RoboDK station: pick and place normal 2r.rdk

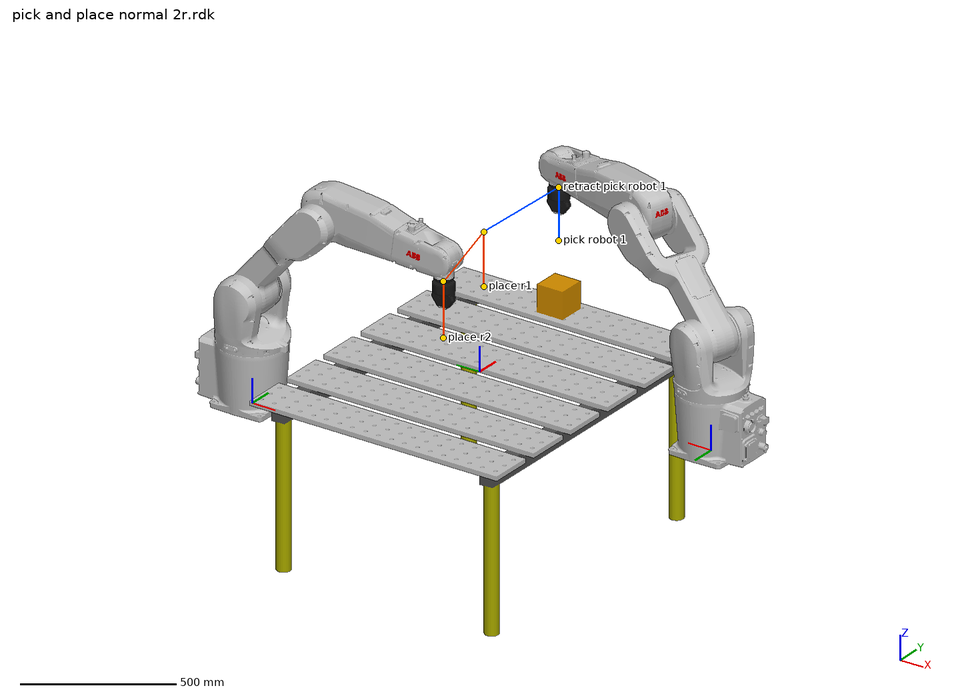
[picture v0: the station drawn from its stored meshes, robots at their saved joint values, targets as dots, program paths as lines]
Station pick and place normal 2r (saved by RoboDK 5.5.0). Poses are relative to the parent item; angles as X-Y-Z fixed-axis rotations.
  - frame Frame 2 at (700, 0, 200) mm, rotated rx 0 ry 0 rz 90 deg
    - object Table 1200x1000mm (Welding) at (0, 0, 0) mm, size 1193.8 x 965.2 x 609.6 mm, geometry from Table-1200x1000mm-Welding.sld
    - object Cube 100mm at (460, 0, 0) mm, size 100 x 100 x 100 mm, geometry from Cube-100mm.sld
  - frame ABB IRB 1200-5/0.9 (1) at (1400, 290, 0) mm, rotated rx 0 ry 0 rz 180 deg
    - robot ABB IRB 1200-5/0.9: 6 axes, payload 5 kg, reach 901 mm, repeatability 0.02 mm, weight 52 kg
        modified DH rows (alpha deg, a mm, theta deg, d mm): 0, 0, 0, 399; -90, 0, -90, 0; 0, 448, 0, 0; -90, 42, 0, 451; 90, 0, 0, 0; -90, 0, 180, 82
        joint limits [-170, -100, -200, -270, -130, -360] to [170, 130, 70, 270, 130, 360]; home [0, 0, 0, 0, 0, 0]; saved at [-16.36, 47.146, -44.021, 0, 86.875, -16.36]
      - robot RobotiQ 2F-140 Gripper (Mechanism) (model RobotiQ 2F140): 1 axes, payload 5 kg
          joint limits [0] to [140]; home [140]; saved at [140]
    - target pick robot 1 (Cartesian target) at (749.42, -220, 449.05) mm, rotated rx 180 ry 0 rz -180 deg; joints [-16.36, 51.781, -27.774, 0, 65.993, -16.36] of ABB IRB 1200-5/0.9
    - target retract pick robot 1 (Cartesian target) at (749.42, -220, 639.05) mm, rotated rx 180 ry 0 rz -180 deg; joints [-16.36, 47.146, -44.021, 0, 86.875, -16.36] of ABB IRB 1200-5/0.9
    - target retract place r1 (Cartesian target) at (759, 184.18, 639.12) mm, rotated rx 180 ry 0.01 rz -179.36 deg; joints [13.64, 47.14, -44.02, 0, 86.87, 13] of ABB IRB 1200-5/0.9
    - target place r1 (Cartesian target) at (759.03, 184.19, 444.12) mm, rotated rx 180 ry 0.01 rz -179.36 deg; joints [13.64, 52.024, -27.559, 0, 65.525, 13] of ABB IRB 1200-5/0.9
  - frame ABB IRB 1200-5/0.9 (2) at (0, -270, 0) mm
    - robot ABB IRB 1200-5/0.9: 6 axes, payload 5 kg, reach 901 mm, repeatability 0.02 mm, weight 52 kg
        modified DH rows (alpha deg, a mm, theta deg, d mm): 0, 0, 0, 399; -90, 0, -90, 0; 0, 448, 0, 0; -90, 42, 0, 451; 90, 0, 0, 0; -90, 0, 180, 82
        joint limits [-170, -100, -200, -270, -130, -360] to [170, 130, 70, 270, 130, 360]; home [0, 0, 0, 0, 0, 0]; saved at [0.38, 40.43, -32.71, 0, 82.29, -180.25]
      - robot RobotiQ 2F-140 Gripper (Mechanism) (model RobotiQ 2F140): 1 axes, payload 5 kg
          joint limits [0] to [140]; home [140]; saved at [140]
    - target retract pick r2 (Cartesian target) at (641, 375.82, 639.12) mm, rotated rx 180 ry 0.01 rz 0.64 deg; joints [13.64, 47.14, -44.02, 0, 86.87, 13] of ABB IRB 1200-5/0.9
    - target pick r2 (Cartesian target) at (640.97, 375.81, 444.12) mm, rotated rx 180 ry 0.01 rz 0.64 deg; joints [13.64, 109.487, -141.8, 0, 122.303, 13] of ABB IRB 1200-5/0.9
    - target retract place r2 (Cartesian target) at (743.06, 4.93, 639.05) mm, rotated rx -180 ry 0.01 rz 0.63 deg; joints [0.38, 40.43, -32.71, 0, 82.29, -180.25] of ABB IRB 1200-5/0.9
    - target place r2 (Cartesian target) at (743.03, 4.93, 439.05) mm, rotated rx -180 ry 0.01 rz 0.63 deg; joints [0.38, 47.164, -18.076, 0, 60.923, -180.25] of ABB IRB 1200-5/0.9
  - program Prog 1 robot 1 (8 instructions, listed below)
  - program Prog 2 robot 2 (7 instructions, listed below)
  - program RESET (1 instructions, listed below)
  - program Pick and Place 2 robots (3 instructions, listed below)
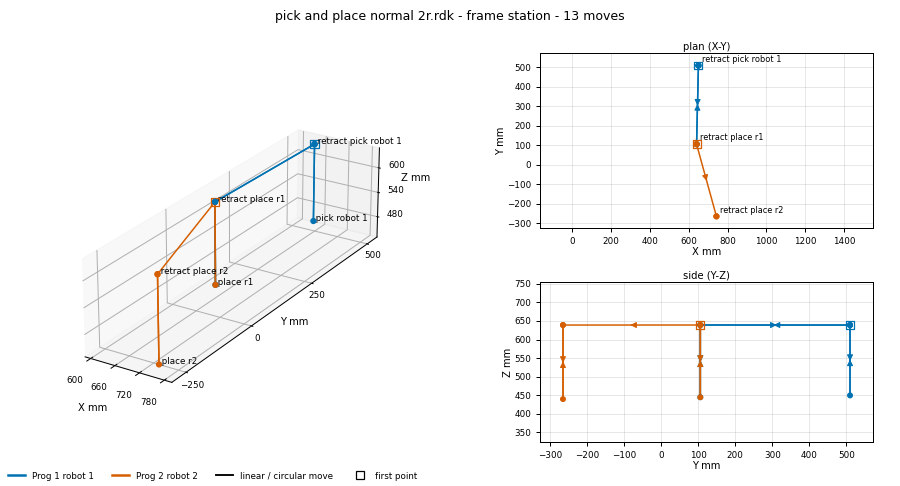
[picture p0: tool path of pick and place normal 2r.rdk in frame station, 13 of 13 moves have a stored position in this frame; points joined in program order, loops and branches not executed]

--- program Prog 1 robot 1 (robot ABB IRB 1200-5/0.9) ---
  Est. Ref.: ABB IRB 1200-5/0.9 (1)
  MoveJ (retract pick robot 1)
  MoveL (pick robot 1)
  MoveL (retract pick robot 1)
  MoveL (retract place r1)
  MoveL (place r1)
  MoveL (retract place r1)
  MoveL (retract pick robot 1)

--- program Prog 2 robot 2 (robot ABB IRB 1200-5/0.9) ---
  Est. Ref.: ABB IRB 1200-5/0.9 (2)
  MoveJ (retract pick r2)
  MoveL (pick r2)
  MoveL (retract pick r2)
  MoveL (retract place r2)
  MoveL (place r2)
  MoveL (retract place r2)

--- program RESET (robot ABB IRB 1200-5/0.9) ---
  Reemplazar Cube 100mm

--- program Pick and Place 2 robots (robot ABB IRB 1200-5/0.9) ---
  Llamar Prog 1 robot 1
  Llamar Prog 2 robot 2
  Llamar RESET
